(* IEC 61131-3 sources: PortalRobot/Portal_robot/Device/application/FB/FB_CELL_MANAGER (part 2) *)

(* ---- FB_CELL_MANAGER.CanReturnHeldBlank.st ---- *)
METHOD PRIVATE CanReturnHeldBlank : BOOL
VAR
	uiMagazine : UINT; // Магазин следующей операции, независимо от магазина возврата
	uiMachine  : UINT;
	uiType     : UINT;
	uiReservedFreeSlots : UINT; // Возврат занимает один универсальный слот своего магазина
END_VAR

// --- BEGIN IMPLEMENTATION ---

CanReturnHeldBlank := FALSE;

// Для одного типа возврат не открывает нового маршрута. Два груза сначала
// разбираются штатным LOAD/PUT; занятый исправный станок своей заготовки ждём.
IF (Config.uiTypeCount > UINT#1)
AND (Config.uiTypeCount <= UINT#3)
AND stRobotStatus.xBlankAvailable
AND NOT stRobotStatus.xDetailAvailable
AND NOT stRobotStatus.xBusy
AND NOT xStopRequested
AND xMagazineReady
AND (uiBlankPayloadType >= UINT#1)
AND (uiBlankPayloadType <= Config.uiTypeCount) THEN
	IF (stMagazineStatus.stTypeStatus.aiFreeSlot[uiBlankPayloadType] > SINT#0)
	AND (SelectMachineForHeldBlank(
		uiProductType := uiBlankPayloadType,
		uiCurrentMachine := uiSelectedMachine
	) = UINT#0) THEN
		FOR uiMagazine := UINT#1 TO GVL_CELL_SETTINGS.MagazineCount DO
			IF ((uiMagazine = UINT#1) AND xMagazine1Available)
			OR ((uiMagazine = UINT#2) AND xMagazine2Available) THEN
				uiReservedFreeSlots := UINT#0;
				IF uiMagazine = uiActiveMagazine THEN
					uiReservedFreeSlots := UINT#1;
				END_IF;
				FOR uiMachine := FIRST_MACHINE TO LAST_MACHINE DO
					IF IsMachineEligible(uiMachine := uiMachine) THEN
						uiType := Config.auiMachineType[uiMachine];
						IF uiType <> uiBlankPayloadType THEN
							// TAKE освобождает место даже в полной палете. Работающий
							// станок другого типа допускает обычное ожидание его цикла.
							IF (astMagazineStatus[uiMagazine].stTypeStatus.aiBlankSlot[uiType] > SINT#0)
							AND (astMachineStatus[uiMachine].xProcessing
								OR axMachineStartPending[uiMachine]
								OR (astMachineStatus[uiMachine].xCanAcceptService
									AND ((astMachineStatus[uiMachine].ePartState = E_PART_STATE.EMPTY)
										OR astMachineStatus[uiMachine].xServiceRequired))) THEN
								CanReturnHeldBlank := TRUE;
							END_IF;
							// Отдельная выгрузка полезна только для уже готовой детали.
							// Последний свободный слот нельзя занять возвратом и затем
							// выдать UNLOAD без места для этой детали.
							IF astMachineStatus[uiMachine].xCanAcceptService
							AND astMachineStatus[uiMachine].xServiceRequired
							AND (astMachineStatus[uiMachine].ePartState = E_PART_STATE.LOADED)
							AND (astMachineStatus[uiMachine].ePartType = E_PART_TYPE.DETAIL)
							AND (astMagazineStatus[uiMagazine].stTypeStatus.auiFreeCount[uiType] > uiReservedFreeSlots) THEN
								CanReturnHeldBlank := TRUE;
							END_IF;
						END_IF;
					END_IF;
				END_FOR;
			END_IF;
		END_FOR;
	END_IF;
END_IF;

(* ---- FB_CELL_MANAGER.HasMagazineWork.st ---- *)
METHOD PRIVATE HasMagazineWork : BOOL
VAR_INPUT
	uiMagazine : UINT; // Оцениваемый магазин; активный владелец не меняется
	xSupplyBlankOnly : BOOL; // TRUE: нужна именно допустимая подача заготовки
END_VAR
VAR
	uiMachine : UINT;
	uiType : UINT;
	xPending : BOOL;
END_VAR

// --- BEGIN IMPLEMENTATION ---

HasMagazineWork := FALSE;
IF (uiMagazine >= UINT#1) AND (uiMagazine <= UINT#2) THEN
	FOR uiMachine := FIRST_MACHINE TO LAST_MACHINE DO
		IF IsMachineEligible(uiMachine := uiMachine) THEN
			uiType := Config.auiMachineType[uiMachine];
			IF (uiType >= UINT#1) AND (uiType <= UINT#3) THEN
				xPending := IsMachineWorkPending(uiMachine := uiMachine);
				// Те же критерии, что у SelectMachineBeforeTake: готовый
				// LOAD/CHANGE либо ожидаемое автоматическое обслуживание.
				IF (astMagazineStatus[uiMagazine].stTypeStatus.aiBlankSlot[uiType] > SINT#0)
				AND (xPending OR (astMachineStatus[uiMachine].xCanAcceptService
					AND ((astMachineStatus[uiMachine].ePartState = E_PART_STATE.EMPTY)
						OR astMachineStatus[uiMachine].xServiceRequired))) THEN
					HasMagazineWork := TRUE;
				END_IF;
				// Без заготовки остаётся отдельный UNLOAD в свободный слот.
				IF NOT xSupplyBlankOnly
				AND (astMagazineStatus[uiMagazine].stTypeStatus.aiFreeSlot[uiType] > SINT#0)
				AND (xPending OR (astMachineStatus[uiMachine].xCanAcceptService
					AND astMachineStatus[uiMachine].xServiceRequired
					AND (astMachineStatus[uiMachine].ePartState = E_PART_STATE.LOADED)
					AND (astMachineStatus[uiMachine].ePartType = E_PART_TYPE.DETAIL))) THEN
					HasMagazineWork := TRUE;
				END_IF;
			END_IF;
		END_IF;
	END_FOR;
END_IF;

(* ---- FB_CELL_MANAGER.IsMachineCompatible.st ---- *)
METHOD PRIVATE IsMachineCompatible : BOOL
VAR_INPUT
	uiMachine     : UINT; // Проверяемый станок
	uiProductType : UINT; // Тип заготовки в захвате
END_VAR

// --- BEGIN IMPLEMENTATION ---

IsMachineCompatible := IsMachineEligible(uiMachine := uiMachine);
IF IsMachineCompatible THEN
	IsMachineCompatible := (uiProductType >= UINT#1)
		AND (uiProductType <= Config.uiTypeCount)
		AND (Config.auiMachineType[uiMachine] = uiProductType);
END_IF;

(* ---- FB_CELL_MANAGER.IsMachineEligible.st ---- *)
METHOD PRIVATE IsMachineEligible : BOOL
VAR_INPUT
	uiMachine : UINT; // Проверяемый станок
END_VAR

// --- BEGIN IMPLEMENTATION ---

IsMachineEligible := (uiMachine >= FIRST_MACHINE)
	AND (uiMachine <= LAST_MACHINE);

IF IsMachineEligible THEN
	IsMachineEligible := astMachineStatus[uiMachine].xEnabled
		AND NOT astMachineStatus[uiMachine].xError
		AND NOT astMachineStatus[uiMachine].xDisablePending
		AND NOT axGeometryUnloadBlocked[uiMachine]
		AND (Config.auiMachineType[uiMachine] >= UINT#1)
		AND (Config.auiMachineType[uiMachine] <= Config.uiTypeCount);
END_IF;

(* ---- FB_CELL_MANAGER.IsMachineWorkPending.st ---- *)
METHOD PRIVATE IsMachineWorkPending : BOOL
VAR_INPUT
	uiMachine : UINT; // Проверяемый станок
END_VAR

// --- BEGIN IMPLEMENTATION ---

IsMachineWorkPending := FALSE;
IF IsMachineEligible(uiMachine := uiMachine) THEN
	// LOADED сам по себе не обещает автоматического продолжения: оператор
	// может ещё не разрешить цикл. Сохраняем обработку, подтверждение запуска
	// и короткий автоматический переход после обработки/обслуживания.
	IsMachineWorkPending := astMachineStatus[uiMachine].xProcessing
		OR axMachineStartPending[uiMachine]
		OR ((astMachineStatus[uiMachine].ePartState = E_PART_STATE.LOADED)
			AND ((astMachineStatus[uiMachine].ePartType = E_PART_TYPE.PART)
				OR (astMachineStatus[uiMachine].ePartType = E_PART_TYPE.DETAIL))
			AND (astMachineStatus[uiMachine].xBusy
				OR astMachineStatus[uiMachine].xDone));
END_IF;

(* ---- FB_CELL_MANAGER.PlanGeometry.st ---- *)
METHOD PRIVATE PlanGeometry : BOOL
VAR
	uiFree : UINT;
	uiAvailable : UINT;
END_VAR

// --- BEGIN IMPLEMENTATION ---

PlanGeometry := FALSE;
IF xGeometryHeld AND stRobotStatus.xDetailAvailable AND (uiGeometryMachine >= UINT#1) AND (uiGeometryMachine <= UINT#3) THEN
	uiFree := F_GEOMETRY_SELECT_STATION(xRequireFree := TRUE, uiMachine := uiGeometryMachine);
	uiAvailable := F_GEOMETRY_SELECT_STATION(xRequireFree := FALSE, uiMachine := uiGeometryMachine);
	IF uiFree > UINT#0 THEN
		uiGeometryStation := uiFree; uiGeometryStep := UINT#0;
		GVL_GEOMETRY_CONTROL.astCalls[uiGeometryMachine].uiStation := uiFree;
		GVL_GEOMETRY_CONTROL.astCalls[uiGeometryMachine].uiState := UINT#3;
		GVL_GEOMETRY_CONTROL.astCalls[uiGeometryMachine].uiReason := UINT#0;
		F_GEOMETRY_EVENT(Call := GVL_GEOMETRY_CONTROL.astCalls[uiGeometryMachine]);
		GVL_GEOMETRY_CONTROL.astSignals[uiFree].Call := GVL_GEOMETRY_CONTROL.astCalls[uiGeometryMachine];
		GVL_GEOMETRY_CONTROL.astSignals[uiFree].xReserve := TRUE;
		eState := E_CELL_MANAGER_STATE.GEOMETRY_DELIVER; PlanGeometry := TRUE;
	ELSIF (uiAvailable > UINT#0) AND Persistent_Value.xWaitWhenOccupied THEN
		uiGeometryParkStation := uiAvailable;
		eState := E_CELL_MANAGER_STATE.GEOMETRY_WAIT_FREE; PlanGeometry := TRUE;
	ELSE
		// Окончательный журнал магазина формируем только по фактической укладке.
		IF uiAvailable > UINT#0 THEN uiGeometryBypassReason := UINT#1; ELSE uiGeometryBypassReason := UINT#2; END_IF;
		udiGeometryMagazineCounter := stMagazineStatus.udiProducedPartsTotal;
	END_IF;
END_IF;

(* ---- FB_CELL_MANAGER.RaisePayloadRouteWarning.st ---- *)
METHOD PRIVATE RaisePayloadRouteWarning
VAR_INPUT
	uiPayloadType     : UINT;
	uiDestinationType : UINT;
END_VAR

// --- BEGIN IMPLEMENTATION ---

IF (uiPayloadType >= UINT#1)
AND (uiDestinationType >= UINT#1)
AND (uiPayloadType <> uiDestinationType) THEN
	IF NOT xPayloadRouteWarningActive THEN
		Diag.stWarning.uiCode := WRN_PAYLOAD_ROUTE_MISMATCH;
		Diag.stWarning.udiSequence := Diag.stWarning.udiSequence + UDINT#1;
		IF Diag.stWarning.udiSequence = UDINT#0 THEN
			Diag.stWarning.udiSequence := UDINT#1;
		END_IF;
		xPayloadRouteWarningActive := TRUE;
	END_IF;
ELSE
	xPayloadRouteWarningActive := FALSE;
END_IF;

(* ---- FB_CELL_MANAGER.RunGeometryRoute.st ---- *)
METHOD PRIVATE RunGeometryRoute

// --- BEGIN IMPLEMENTATION ---

CASE eState OF
	E_CELL_MANAGER_STATE.GEOMETRY_WAIT_FREE:
		IF uiGeometryParkStation = UINT#1 THEN eGeometrySafePoint := E_POINT_NAME.GEOMETRY_1_SAFE;
		ELSE eGeometrySafePoint := E_POINT_NAME.GEOMETRY_2_SAFE; END_IF;
		IF stRobotStatus.xBusy OR stRobotStatus.xDone OR xMotionBusy THEN
			// Освобождение ГК не отменяет уже выданное парковочное движение.
			Command.stRobot.xExecute := TRUE; Command.stRobot.eAction := E_ROBOT_ACTION.MOVE_TO_POINT;
			Command.stRobot.eSetPoint := eGeometrySafePoint;
			IF stRobotStatus.xDone THEN eGeometryReturnState := E_CELL_MANAGER_STATE.GEOMETRY_WAIT_FREE; eState := E_CELL_MANAGER_STATE.GEOMETRY_RELEASE_COMMAND; END_IF;
		ELSIF xStopRequested THEN
			xRunning := FALSE; eState := E_CELL_MANAGER_STATE.IDLE;
		ELSIF F_GEOMETRY_SELECT_STATION(xRequireFree := TRUE, uiMachine := uiGeometryMachine) > UINT#0 THEN
			eState := E_CELL_MANAGER_STATE.PLAN_TARGET;
		ELSIF (F_GEOMETRY_SELECT_STATION(xRequireFree := FALSE, uiMachine := uiGeometryMachine) = UINT#0) OR NOT Persistent_Value.xWaitWhenOccupied THEN
			eState := E_CELL_MANAGER_STATE.PLAN_TARGET;
		ELSE
			// Ожидаем с деталью в захвате на безопасной высоте; конвейер может работать.
			IF uiGeometryParkStation = UINT#1 THEN eGeometrySafePoint := E_POINT_NAME.GEOMETRY_1_SAFE;
			ELSE eGeometrySafePoint := E_POINT_NAME.GEOMETRY_2_SAFE; END_IF;
			IF stRobotStatus.eCurrentPoint <> eGeometrySafePoint THEN
				Command.stRobot.xExecute := TRUE; Command.stRobot.eAction := E_ROBOT_ACTION.MOVE_TO_POINT;
				Command.stRobot.eSetPoint := eGeometrySafePoint;
				IF stRobotStatus.xDone THEN eGeometryReturnState := E_CELL_MANAGER_STATE.GEOMETRY_WAIT_FREE; eState := E_CELL_MANAGER_STATE.GEOMETRY_RELEASE_COMMAND; END_IF;
			END_IF;
		END_IF;
	E_CELL_MANAGER_STATE.GEOMETRY_DELIVER:
		IF (uiGeometryStation < UINT#1) OR (uiGeometryStation > UINT#2) THEN
			Error.dwErrorActive := Error.dwErrorActive OR ERR_ROBOT; eState := E_CELL_MANAGER_STATE.ERROR;
		ELSIF GVL_GEOMETRY_CONTROL.astStatus[uiGeometryStation].xError
		AND NOT GVL_GEOMETRY_CONTROL.astSignals[uiGeometryStation].xRobotInteraction THEN
			// Оборудование отказало до входа: робот может выбрать другой ГК.
			GVL_GEOMETRY_CONTROL.astSignals[uiGeometryStation].xReserve := FALSE;
			GVL_GEOMETRY_CONTROL.astSignals[uiGeometryStation].xReleased := TRUE;
			GVL_GEOMETRY_CONTROL.astCalls[uiGeometryMachine].uiStation := UINT#0;
			GVL_GEOMETRY_CONTROL.astCalls[uiGeometryMachine].uiState := UINT#2;
			GVL_GEOMETRY_CONTROL.astCalls[uiGeometryMachine].uiReason := UINT#4;
			F_GEOMETRY_EVENT(Call := GVL_GEOMETRY_CONTROL.astCalls[uiGeometryMachine]);
			uiGeometryStation := UINT#0; eState := E_CELL_MANAGER_STATE.PLAN_TARGET;
		ELSIF NOT GVL_GEOMETRY_CONTROL.astSignals[uiGeometryStation].xRobotInteraction
		AND (NOT GVL_GEOMETRY_CONTROL.astStatus[uiGeometryStation].xEnabled
			OR (GVL_GEOMETRY_CONTROL.astStatus[uiGeometryStation].uiState = UINT#5)
			OR GVL_GEOMETRY_CONTROL.astStatus[uiGeometryStation].xDriveRunning) THEN
			// Выключение в том же скане, что резерв, не разрешает вход робота.
			GVL_GEOMETRY_CONTROL.astSignals[uiGeometryStation].xReserve := FALSE;
			GVL_GEOMETRY_CONTROL.astSignals[uiGeometryStation].xReleased := TRUE;
			GVL_GEOMETRY_CONTROL.astCalls[uiGeometryMachine].uiStation := UINT#0;
			GVL_GEOMETRY_CONTROL.astCalls[uiGeometryMachine].uiState := UINT#2;
			GVL_GEOMETRY_CONTROL.astCalls[uiGeometryMachine].uiReason := UINT#3;
			F_GEOMETRY_EVENT(Call := GVL_GEOMETRY_CONTROL.astCalls[uiGeometryMachine]);
			uiGeometryStation := UINT#0; eState := E_CELL_MANAGER_STATE.PLAN_TARGET;
		ELSIF GVL_GEOMETRY_CONTROL.astStatus[uiGeometryStation].xError OR stRobotStatus.xError OR xGlobalError THEN
			xSafetyHomeRequired := TRUE; xStoppedPoseValid := FALSE;
			Error.dwErrorActive := Error.dwErrorActive OR ERR_ROBOT; eState := E_CELL_MANAGER_STATE.ERROR;
		ELSIF GVL_GEOMETRY_CONTROL.astStatus[uiGeometryStation].xReserved THEN
			IF uiGeometryStation = UINT#1 THEN
				eGeometrySafePoint := E_POINT_NAME.GEOMETRY_1_SAFE; eGeometryPlacePoint := E_POINT_NAME.GEOMETRY_1_PLACE;
			ELSE
				eGeometrySafePoint := E_POINT_NAME.GEOMETRY_2_SAFE; eGeometryPlacePoint := E_POINT_NAME.GEOMETRY_2_PLACE;
			END_IF;
			GVL_GEOMETRY_CONTROL.astSignals[uiGeometryStation].xRobotInteraction := TRUE;
			IF uiGeometryStep <= UINT#4 THEN
				Command.stRobot.xExecute := TRUE; Command.stRobot.eAction := E_ROBOT_ACTION.MOVE_TO_POINT;
				CASE uiGeometryStep OF
					UINT#0, UINT#4: Command.stRobot.eSetPoint := eGeometrySafePoint;
					// Для укладки на ГК нужна ориентация «к заготовке»; поворот выполняется на SAFE.
					UINT#1: Command.stRobot.eAction := E_ROBOT_ACTION.ROTATE_TO_BLANK;
					UINT#2: Command.stRobot.eSetPoint := eGeometryPlacePoint;
					UINT#3: Command.stRobot.eAction := E_ROBOT_ACTION.UNCLAMP_2;
				END_CASE;
				IF stRobotStatus.xDone THEN
					IF uiGeometryStep = UINT#3 THEN
						IF stRobotStatus.xGripper2Open AND NOT stRobotStatus.xDetailAvailable THEN
							GVL_GEOMETRY_CONTROL.astSignals[uiGeometryStation].xDeposited := TRUE;
							uiDetailPayloadType := UINT#0;
						ELSE Error.dwErrorActive := Error.dwErrorActive OR ERR_ROBOT; eState := E_CELL_MANAGER_STATE.ERROR; END_IF;
					END_IF;
					IF eState <> E_CELL_MANAGER_STATE.ERROR THEN
						eGeometryReturnState := E_CELL_MANAGER_STATE.GEOMETRY_DELIVER;
						eState := E_CELL_MANAGER_STATE.GEOMETRY_RELEASE_COMMAND;
					END_IF;
				END_IF;
			ELSE
				GVL_GEOMETRY_CONTROL.astSignals[uiGeometryStation].xReserve := FALSE;
				GVL_GEOMETRY_CONTROL.astSignals[uiGeometryStation].xDeposited := FALSE;
				GVL_GEOMETRY_CONTROL.astSignals[uiGeometryStation].xRobotInteraction := FALSE;
				GVL_GEOMETRY_CONTROL.astSignals[uiGeometryStation].xReleased := TRUE;
				GVL_GEOMETRY_CONTROL.uiLastStation := uiGeometryStation;
				xGeometryHeld := FALSE; uiGeometryMachine := UINT#0; uiGeometryStation := UINT#0;
				eState := E_CELL_MANAGER_STATE.PLAN_TARGET;
			END_IF;
		ELSE
			// Потеря резерва в зоне робота требует восстановления, а не нового маршрута.
			IF GVL_GEOMETRY_CONTROL.astSignals[uiGeometryStation].xRobotInteraction THEN
				xSafetyHomeRequired := TRUE; xStoppedPoseValid := FALSE;
				Error.dwErrorActive := Error.dwErrorActive OR ERR_ROBOT; eState := E_CELL_MANAGER_STATE.ERROR;
			ELSIF NOT GVL_GEOMETRY_CONTROL.astStatus[uiGeometryStation].xReady
			OR (GVL_GEOMETRY_CONTROL.astStatus[uiGeometryStation].uiState = UINT#5) THEN
				GVL_GEOMETRY_CONTROL.astSignals[uiGeometryStation].xReserve := FALSE;
				GVL_GEOMETRY_CONTROL.astSignals[uiGeometryStation].xReleased := TRUE;
				GVL_GEOMETRY_CONTROL.astCalls[uiGeometryMachine].uiStation := UINT#0;
				GVL_GEOMETRY_CONTROL.astCalls[uiGeometryMachine].uiState := UINT#2;
				GVL_GEOMETRY_CONTROL.astCalls[uiGeometryMachine].uiReason := UINT#3;
				F_GEOMETRY_EVENT(Call := GVL_GEOMETRY_CONTROL.astCalls[uiGeometryMachine]);
				uiGeometryStation := UINT#0; eState := E_CELL_MANAGER_STATE.PLAN_TARGET;
			END_IF;
		END_IF;
	E_CELL_MANAGER_STATE.GEOMETRY_RELEASE_COMMAND:
		IF stRobotStatus.xError THEN
			xSafetyHomeRequired := TRUE; xStoppedPoseValid := FALSE;
			Error.dwErrorActive := Error.dwErrorActive OR ERR_ROBOT; eState := E_CELL_MANAGER_STATE.ERROR;
		ELSIF NOT stRobotStatus.xBusy AND NOT stRobotStatus.xDone THEN
			IF eGeometryReturnState = E_CELL_MANAGER_STATE.GEOMETRY_DELIVER THEN uiGeometryStep := uiGeometryStep + UINT#1; END_IF;
			eState := eGeometryReturnState;
		END_IF;
END_CASE;

(* ---- FB_CELL_MANAGER.SelectMachineBeforeTake.st ---- *)
METHOD PRIVATE SelectMachineBeforeTake : UINT
VAR
	uiMachine           : UINT; // Проверяемый станок
	uiType              : UINT; // Тип станка
	xTimedFound         : BOOL; // Найден кандидат с оценкой времени
	tMinimumRemaining   : TIME; // Минимальное найденное оставшееся время
	tCandidateRemaining : TIME; // Оценка кандидата, который подтверждает запуск цикла
END_VAR

// --- BEGIN IMPLEMENTATION ---

SelectMachineBeforeTake := UINT#0;
xTimedFound := FALSE;
tMinimumRemaining := T#0S;

// Сначала выбирается станок, который можно обслужить без ожидания.
// xPartReady отдельно не используется: после завершения обслуживания он может
// сохраняться до перехода FB_MACHINE из DONE в IDLE и повторно выбрать тот же станок.
FOR uiMachine := FIRST_MACHINE TO LAST_MACHINE DO
	uiType := Config.auiMachineType[uiMachine];
	IF IsMachineEligible(uiMachine := uiMachine) THEN
		IF (SelectMachineBeforeTake = UINT#0)
		AND (stMagazineStatus.stTypeStatus.aiBlankSlot[uiType] > SINT#0)
		AND astMachineStatus[uiMachine].xCanAcceptService
		AND ((astMachineStatus[uiMachine].ePartState = E_PART_STATE.EMPTY)
			OR astMachineStatus[uiMachine].xServiceRequired) THEN
			SelectMachineBeforeTake := uiMachine;
		END_IF;
	END_IF;
END_FOR;

// Затем сравниваются фактически обрабатывающие станки по оставшемуся времени.
IF SelectMachineBeforeTake = UINT#0 THEN
	FOR uiMachine := FIRST_MACHINE TO LAST_MACHINE DO
		uiType := Config.auiMachineType[uiMachine];
		IF IsMachineEligible(uiMachine := uiMachine) THEN
			IF (stMagazineStatus.stTypeStatus.aiBlankSlot[uiType] > SINT#0)
			AND astMachineStatus[uiMachine].xProcessing
			AND astMachineStatus[uiMachine].xCycleTimeValid THEN
				IF NOT xTimedFound
				OR (astMachineStatus[uiMachine].tRemaining < tMinimumRemaining) THEN
					SelectMachineBeforeTake := uiMachine;
					tMinimumRemaining := astMachineStatus[uiMachine].tRemaining;
					xTimedFound := TRUE;
				END_IF;
			END_IF;
		END_IF;
	END_FOR;
END_IF;

// Только что обслуженный станок может появиться в xProcessing на несколько циклов PLC позже.
// До подтверждения запуска он участвует в том же сравнении по полному tCycleExpected.
IF (SelectMachineBeforeTake = UINT#0) OR xTimedFound THEN
	FOR uiMachine := FIRST_MACHINE TO LAST_MACHINE DO
		uiType := Config.auiMachineType[uiMachine];
		IF axMachineStartPending[uiMachine]
		AND IsMachineEligible(uiMachine := uiMachine)
		AND (stMagazineStatus.stTypeStatus.aiBlankSlot[uiType] > SINT#0)
		AND astMachineStatus[uiMachine].xCycleTimeValid THEN
			tCandidateRemaining := START_PENDING_ESTIMATE
				+ astMachineStatus[uiMachine].tCycleExpected;
			IF NOT xTimedFound
			OR (tCandidateRemaining < tMinimumRemaining) THEN
				SelectMachineBeforeTake := uiMachine;
				tMinimumRemaining := tCandidateRemaining;
				xTimedFound := TRUE;
			END_IF;
		END_IF;
	END_FOR;
END_IF;

// Неизвестное время не делает включённый исправный станок недоступным.
IF (SelectMachineBeforeTake = UINT#0) AND NOT xTimedFound THEN
	FOR uiMachine := FIRST_MACHINE TO LAST_MACHINE DO
		uiType := Config.auiMachineType[uiMachine];
		IF IsMachineEligible(uiMachine := uiMachine) THEN
			IF (SelectMachineBeforeTake = UINT#0)
			AND (stMagazineStatus.stTypeStatus.aiBlankSlot[uiType] > SINT#0)
			AND IsMachineWorkPending(uiMachine := uiMachine) THEN
				SelectMachineBeforeTake := uiMachine;
			END_IF;
		END_IF;
	END_FOR;
END_IF;

(* ---- FB_CELL_MANAGER.SelectMachineForHeldBlank.st ---- *)
METHOD PRIVATE SelectMachineForHeldBlank : UINT
VAR_INPUT
	uiProductType    : UINT; // Тип уже взятой заготовки
	uiCurrentMachine : UINT; // Текущая цель для устойчивого повторного выбора
END_VAR
VAR
	uiMachine           : UINT; // Проверяемый станок
	xTimedFound         : BOOL; // Найден станок с оценкой времени
	xCurrentTimed       : BOOL; // Текущая цель имеет сопоставимую оценку
	tMinimumRemaining   : TIME; // Минимальное оставшееся время
	tCandidateRemaining : TIME; // Оценка проверяемого станка
	tCurrentRemaining   : TIME; // Оценка текущей цели
END_VAR

// --- BEGIN IMPLEMENTATION ---

SelectMachineForHeldBlank := UINT#0;
xTimedFound := FALSE;
xCurrentTimed := FALSE;
tMinimumRemaining := T#0S;
tCandidateRemaining := T#0S;
tCurrentRemaining := T#0S;

// UINT#0 означает, что после остановки/аварии текущая цель ещё не выбрана.
// Проверка диапазона вынесена отдельно: обычный AND в CODESYS вычисляет все
// операнды и не защищает ARRAY [1..3] от обращения по индексу 0.
IF (uiCurrentMachine >= FIRST_MACHINE)
AND (uiCurrentMachine <= LAST_MACHINE) THEN
	// Если робот уже находится у готовой совместимой цели, лишнее перемещение не требуется.
	IF IsMachineCompatible(
		uiMachine := uiCurrentMachine,
		uiProductType := uiProductType
	)
	AND astMachineStatus[uiCurrentMachine].xCanAcceptService
	AND ((astMachineStatus[uiCurrentMachine].ePartState = E_PART_STATE.EMPTY)
		OR astMachineStatus[uiCurrentMachine].xServiceRequired) THEN
		SelectMachineForHeldBlank := uiCurrentMachine;
	END_IF;
END_IF;

// Готовая совместимая цель имеет приоритет. Переходный xPartReady без
// xCanAcceptService не считается разрешением на повторное обслуживание.
FOR uiMachine := FIRST_MACHINE TO LAST_MACHINE DO
	IF (SelectMachineForHeldBlank = UINT#0)
	AND IsMachineEligible(uiMachine := uiMachine)
	AND (Config.auiMachineType[uiMachine] = uiProductType)
	AND astMachineStatus[uiMachine].xCanAcceptService
	AND ((astMachineStatus[uiMachine].ePartState = E_PART_STATE.EMPTY)
		OR astMachineStatus[uiMachine].xServiceRequired) THEN
		SelectMachineForHeldBlank := uiMachine;
	END_IF;
END_FOR;

// Обрабатывающие и только что запущенные совместимые станки сравниваются
// по одному прогнозу: tRemaining либо полный tCycleExpected для start-pending.
IF SelectMachineForHeldBlank = UINT#0 THEN
	FOR uiMachine := FIRST_MACHINE TO LAST_MACHINE DO
		IF IsMachineEligible(uiMachine := uiMachine)
		AND (Config.auiMachineType[uiMachine] = uiProductType)
		AND astMachineStatus[uiMachine].xCycleTimeValid THEN
			IF astMachineStatus[uiMachine].xProcessing THEN
				tCandidateRemaining := astMachineStatus[uiMachine].tRemaining;
			ELSIF axMachineStartPending[uiMachine] THEN
				tCandidateRemaining := START_PENDING_ESTIMATE
					+ astMachineStatus[uiMachine].tCycleExpected;
			ELSE
				tCandidateRemaining := T#0S;
			END_IF;

			IF astMachineStatus[uiMachine].xProcessing
			OR axMachineStartPending[uiMachine] THEN
				IF NOT xTimedFound
				OR (tCandidateRemaining < tMinimumRemaining) THEN
					SelectMachineForHeldBlank := uiMachine;
					tMinimumRemaining := tCandidateRemaining;
					xTimedFound := TRUE;
				END_IF;
			END_IF;
		END_IF;
	END_FOR;

	// При почти одинаковом времени сохраняется текущая цель.
	IF xTimedFound
	AND (uiCurrentMachine >= FIRST_MACHINE)
	AND (uiCurrentMachine <= LAST_MACHINE) THEN
		IF (SelectMachineForHeldBlank <> uiCurrentMachine)
		AND IsMachineCompatible(
			uiMachine := uiCurrentMachine,
			uiProductType := uiProductType
		)
		AND astMachineStatus[uiCurrentMachine].xCycleTimeValid THEN
			xCurrentTimed := astMachineStatus[uiCurrentMachine].xProcessing
				OR axMachineStartPending[uiCurrentMachine];
			IF astMachineStatus[uiCurrentMachine].xProcessing THEN
				tCurrentRemaining := astMachineStatus[uiCurrentMachine].tRemaining;
			ELSIF axMachineStartPending[uiCurrentMachine] THEN
				tCurrentRemaining := START_PENDING_ESTIMATE
					+ astMachineStatus[uiCurrentMachine].tCycleExpected;
			END_IF;
			IF xCurrentTimed
			AND (tCurrentRemaining >= tMinimumRemaining)
			AND ((tCurrentRemaining - tMinimumRemaining) <= MACHINE_SWITCH_DEADBAND) THEN
				SelectMachineForHeldBlank := uiCurrentMachine;
			END_IF;
		END_IF;
	END_IF;
END_IF;

// Без точной оценки сохраняется текущий обрабатывающий маршрут либо выбирается
// первый совместимый обрабатывающий/start-pending станок.
IF SelectMachineForHeldBlank = UINT#0 THEN
	IF (uiCurrentMachine >= FIRST_MACHINE)
	AND (uiCurrentMachine <= LAST_MACHINE) THEN
		IF IsMachineCompatible(
			uiMachine := uiCurrentMachine,
			uiProductType := uiProductType
		)
		AND (astMachineStatus[uiCurrentMachine].xProcessing
			OR axMachineStartPending[uiCurrentMachine]) THEN
			SelectMachineForHeldBlank := uiCurrentMachine;
		END_IF;
	END_IF;

	FOR uiMachine := FIRST_MACHINE TO LAST_MACHINE DO
		IF (SelectMachineForHeldBlank = UINT#0)
		AND IsMachineEligible(uiMachine := uiMachine)
		AND (Config.auiMachineType[uiMachine] = uiProductType)
		AND (astMachineStatus[uiMachine].xProcessing
			OR axMachineStartPending[uiMachine]) THEN
			SelectMachineForHeldBlank := uiMachine;
		END_IF;
	END_FOR;
END_IF;

// Включённая исправная цель сохраняет ожидание своей заготовки, даже если
// станок ещё не готов. Нулевой результат только разрешает проверку полезности
// возврата в SELECT_FALLBACK; сам по себе он не требует RETURN_BLANK.
IF SelectMachineForHeldBlank = UINT#0 THEN
	IF (uiCurrentMachine >= FIRST_MACHINE)
	AND (uiCurrentMachine <= LAST_MACHINE) THEN
		IF IsMachineCompatible(
			uiMachine := uiCurrentMachine,
			uiProductType := uiProductType
		) THEN
			SelectMachineForHeldBlank := uiCurrentMachine;
		END_IF;
	END_IF;

	FOR uiMachine := FIRST_MACHINE TO LAST_MACHINE DO
		IF (SelectMachineForHeldBlank = UINT#0)
		AND IsMachineEligible(uiMachine := uiMachine)
		AND (Config.auiMachineType[uiMachine] = uiProductType) THEN
			SelectMachineForHeldBlank := uiMachine;
		END_IF;
	END_FOR;
END_IF;

(* ---- FB_CELL_MANAGER.SelectMachineForUnload.st ---- *)
METHOD PRIVATE SelectMachineForUnload : UINT
VAR_INPUT
	uiCurrentMachine : UINT; // Текущая цель для устойчивого повторного выбора
END_VAR
VAR
	uiMachine           : UINT; // Проверяемый станок
	uiType              : UINT; // Тип детали станка
	xTimedFound         : BOOL; // Найден станок с оценкой времени
	xCurrentTimed       : BOOL; // Текущая цель имеет сопоставимую оценку
	tMinimumRemaining   : TIME; // Минимальное найденное оставшееся время
	tCandidateRemaining : TIME; // Оценка проверяемого станка
	tCurrentRemaining   : TIME; // Оценка текущей цели
END_VAR

// --- BEGIN IMPLEMENTATION ---

SelectMachineForUnload := UINT#0;
xTimedFound := FALSE;
xCurrentTimed := FALSE;
tMinimumRemaining := T#0S;
tCandidateRemaining := T#0S;
tCurrentRemaining := T#0S;

// Если робот уже ждёт над готовым станком, лишнее перемещение не требуется.
IF (uiCurrentMachine >= FIRST_MACHINE)
AND (uiCurrentMachine <= LAST_MACHINE) THEN
	IF IsMachineEligible(uiMachine := uiCurrentMachine) THEN
		uiType := Config.auiMachineType[uiCurrentMachine];
		IF (stMagazineStatus.stTypeStatus.aiFreeSlot[uiType] > SINT#0)
		AND astMachineStatus[uiCurrentMachine].xCanAcceptService
		AND astMachineStatus[uiCurrentMachine].xServiceRequired
		AND (astMachineStatus[uiCurrentMachine].ePartState = E_PART_STATE.LOADED)
		AND (astMachineStatus[uiCurrentMachine].ePartType = E_PART_TYPE.DETAIL) THEN
			SelectMachineForUnload := uiCurrentMachine;
		END_IF;
	END_IF;
END_IF;

// Готовая деталь имеет приоритет над ожиданием обработки.
FOR uiMachine := FIRST_MACHINE TO LAST_MACHINE DO
	uiType := Config.auiMachineType[uiMachine];
	IF IsMachineEligible(uiMachine := uiMachine) THEN
		IF (SelectMachineForUnload = UINT#0)
		AND astMachineStatus[uiMachine].xCanAcceptService
		AND astMachineStatus[uiMachine].xServiceRequired
		AND (astMachineStatus[uiMachine].ePartState = E_PART_STATE.LOADED)
		AND (astMachineStatus[uiMachine].ePartType = E_PART_TYPE.DETAIL)
		AND (stMagazineStatus.stTypeStatus.aiFreeSlot[uiType] > SINT#0) THEN
			SelectMachineForUnload := uiMachine;
		END_IF;
	END_IF;
END_FOR;

// Если готовых деталей пока нет, робот заранее направляется к станку с
// минимальным оставшимся временем обработки.
IF SelectMachineForUnload = UINT#0 THEN
	FOR uiMachine := FIRST_MACHINE TO LAST_MACHINE DO
		uiType := Config.auiMachineType[uiMachine];
		IF IsMachineEligible(uiMachine := uiMachine) THEN
			IF (stMagazineStatus.stTypeStatus.aiFreeSlot[uiType] > SINT#0)
			AND astMachineStatus[uiMachine].xCycleTimeValid THEN
				IF astMachineStatus[uiMachine].xProcessing THEN
					tCandidateRemaining := astMachineStatus[uiMachine].tRemaining;
				ELSIF axMachineStartPending[uiMachine] THEN
					tCandidateRemaining := START_PENDING_ESTIMATE
						+ astMachineStatus[uiMachine].tCycleExpected;
				ELSE
					tCandidateRemaining := T#0S;
				END_IF;

				IF astMachineStatus[uiMachine].xProcessing
				OR axMachineStartPending[uiMachine] THEN
					IF NOT xTimedFound
					OR (tCandidateRemaining < tMinimumRemaining) THEN
						SelectMachineForUnload := uiMachine;
						tMinimumRemaining := tCandidateRemaining;
						xTimedFound := TRUE;
					END_IF;
				END_IF;
			END_IF;
		END_IF;
	END_FOR;

	// При почти одинаковом времени сохраняется уже выбранная цель.
	IF xTimedFound
	AND (uiCurrentMachine >= FIRST_MACHINE)
	AND (uiCurrentMachine <= LAST_MACHINE) THEN
		IF (SelectMachineForUnload <> uiCurrentMachine)
		AND IsMachineEligible(uiMachine := uiCurrentMachine) THEN
			uiType := Config.auiMachineType[uiCurrentMachine];
			IF (stMagazineStatus.stTypeStatus.aiFreeSlot[uiType] > SINT#0)
			AND astMachineStatus[uiCurrentMachine].xCycleTimeValid THEN
				xCurrentTimed := astMachineStatus[uiCurrentMachine].xProcessing
					OR axMachineStartPending[uiCurrentMachine];
				IF astMachineStatus[uiCurrentMachine].xProcessing THEN
					tCurrentRemaining := astMachineStatus[uiCurrentMachine].tRemaining;
				ELSIF axMachineStartPending[uiCurrentMachine] THEN
					tCurrentRemaining := START_PENDING_ESTIMATE
						+ astMachineStatus[uiCurrentMachine].tCycleExpected;
				END_IF;
				IF xCurrentTimed
				AND (tCurrentRemaining >= tMinimumRemaining)
				AND ((tCurrentRemaining - tMinimumRemaining) <= MACHINE_SWITCH_DEADBAND) THEN
					SelectMachineForUnload := uiCurrentMachine;
				END_IF;
			END_IF;
		END_IF;
	END_IF;
END_IF;

// При неизвестном времени сохраняется текущая цель либо выбирается первый
// обрабатывающийся/только что запущенный станок с доступным слотом.
IF SelectMachineForUnload = UINT#0 THEN
	IF (uiCurrentMachine >= FIRST_MACHINE)
	AND (uiCurrentMachine <= LAST_MACHINE) THEN
		IF IsMachineEligible(uiMachine := uiCurrentMachine) THEN
			uiType := Config.auiMachineType[uiCurrentMachine];
			IF (stMagazineStatus.stTypeStatus.aiFreeSlot[uiType] > SINT#0)
			AND (astMachineStatus[uiCurrentMachine].xProcessing
				OR axMachineStartPending[uiCurrentMachine]) THEN
				SelectMachineForUnload := uiCurrentMachine;
			END_IF;
		END_IF;
	END_IF;

	FOR uiMachine := FIRST_MACHINE TO LAST_MACHINE DO
		uiType := Config.auiMachineType[uiMachine];
		IF IsMachineEligible(uiMachine := uiMachine) THEN
			IF (SelectMachineForUnload = UINT#0)
			AND (stMagazineStatus.stTypeStatus.aiFreeSlot[uiType] > SINT#0)
			AND (astMachineStatus[uiMachine].xProcessing
				OR axMachineStartPending[uiMachine]) THEN
				SelectMachineForUnload := uiMachine;
			END_IF;
		END_IF;
	END_FOR;
END_IF;

// Переход от окончания цикла к готовности двери может занять несколько сканов.
// В это время сохраняется автоматически продолжающий работу станок.
// Ожидание решения оператора при LOADED сюда не входит.
IF SelectMachineForUnload = UINT#0 THEN
	IF (uiCurrentMachine >= FIRST_MACHINE)
	AND (uiCurrentMachine <= LAST_MACHINE) THEN
		IF IsMachineEligible(uiMachine := uiCurrentMachine) THEN
			uiType := Config.auiMachineType[uiCurrentMachine];
			IF (stMagazineStatus.stTypeStatus.aiFreeSlot[uiType] > SINT#0)
			AND IsMachineWorkPending(uiMachine := uiCurrentMachine) THEN
				SelectMachineForUnload := uiCurrentMachine;
			END_IF;
		END_IF;
	END_IF;

	FOR uiMachine := FIRST_MACHINE TO LAST_MACHINE DO
		uiType := Config.auiMachineType[uiMachine];
		IF IsMachineEligible(uiMachine := uiMachine) THEN
			IF (SelectMachineForUnload = UINT#0)
			AND (stMagazineStatus.stTypeStatus.aiFreeSlot[uiType] > SINT#0)
			AND IsMachineWorkPending(uiMachine := uiMachine) THEN
				SelectMachineForUnload := uiMachine;
			END_IF;
		END_IF;
	END_FOR;
END_IF;

(* ---- FB_CELL_MANAGER.UpdateErrorView.st ---- *)
METHOD PRIVATE UpdateErrorView : ST_CELL_ERROR
VAR_INPUT
	dwError : DWORD; // Битовая маска ошибок нового менеджера
END_VAR
VAR
	stError : ST_CELL_ERROR; // Совместимое представление ошибок
END_VAR

// --- BEGIN IMPLEMENTATION ---

stError.BOTH_GRIPPERS_OCCUPIED := (dwError AND ERR_BOTH_GRIPPERS) <> DWORD#0;
stError.ROBOT_ERROR := (dwError AND ERR_ROBOT) <> DWORD#0;
stError.MAGAZINE_ERROR := (dwError AND ERR_MAGAZINE) <> DWORD#0;
stError.MACHINE_ERROR := (dwError AND ERR_MACHINE) <> DWORD#0;
stError.GLOBAL_STOP := (dwError AND ERR_GLOBAL_STOP) <> DWORD#0;
UpdateErrorView := stError;

(* ---- FB_CELL_MANAGER.UpdateGeometryWait.st ---- *)
METHOD PRIVATE UpdateGeometryWait
VAR
	uiMachine : UINT;
	uiFreeStation : UINT;
	uiCallState : UINT;
	xCalled : BOOL;
	xReadyDetail : BOOL;
	xWaiting : BOOL;
	xRaiseWarning : BOOL;
	Call : ST_GEOMETRY_CALL;
	EmptyCall : ST_GEOMETRY_CALL;
END_VAR

// --- BEGIN IMPLEMENTATION ---

uiFreeStation := F_GEOMETRY_SELECT_STATION(xRequireFree := TRUE, uiMachine := UINT#0);
xRaiseWarning := FALSE;
FOR uiMachine := FIRST_MACHINE TO LAST_MACHINE DO
	uiCallState := GVL_GEOMETRY_CONTROL.astCalls[uiMachine].uiState;
	xCalled := uiCallState = UINT#1;
	// Автовызов известен до выгрузки; счётчик меняется только при фактическом взятии.
	IF ((uiCallState = UINT#0) OR (uiCallState > UINT#3))
	AND GVL_GEOMETRY_CONTROL.xSupported AND Persistent_Value.xAutoEnabled
	AND (GVL_GEOMETRY_CONTROL.astStatus[1].xEnabled OR GVL_GEOMETRY_CONTROL.astStatus[2].xEnabled)
	AND (GVL_GEOMETRY_CONTROL.auiActiveCount[uiMachine] >= (MAX(UINT#1, Persistent_Value.auiPeriod[uiMachine]) - UINT#1)) THEN
		xCalled := TRUE;
	END_IF;
	xReadyDetail := astMachineStatus[uiMachine].xEnabled
		AND NOT astMachineStatus[uiMachine].xError AND NOT astMachineStatus[uiMachine].xDisablePending
		AND NOT astMachineStatus[uiMachine].xBusy AND NOT astMachineStatus[uiMachine].xProcessing
		AND astMachineStatus[uiMachine].xCanAcceptService AND astMachineStatus[uiMachine].xServiceRequired
		AND (astMachineStatus[uiMachine].ePartState = E_PART_STATE.LOADED)
		AND (astMachineStatus[uiMachine].ePartType = E_PART_TYPE.DETAIL);
	IF xRunning AND NOT xManual AND xCalled AND xReadyDetail AND (uiCallState <> UINT#1) THEN
		Persistent_Value.udiNextCallId := Persistent_Value.udiNextCallId + UDINT#1;
		IF Persistent_Value.udiNextCallId = UDINT#0 THEN Persistent_Value.udiNextCallId := UDINT#1; END_IF;
		Call := EmptyCall; Call.udiId := Persistent_Value.udiNextCallId;
		Call.uiMachine := uiMachine; Call.uiProductType := Config.auiMachineType[uiMachine]; Call.uiState := UINT#1;
		GVL_GEOMETRY_CONTROL.astCalls[uiMachine] := Call;
		F_GEOMETRY_EVENT(Call := Call);
	END_IF;
	// Пустой станок можно загрузить. Уже начатый рецепт не прерываем.
	axGeometryUnloadBlocked[uiMachine] := xCalled AND (uiFreeStation = UINT#0)
		AND (astMachineStatus[uiMachine].ePartState = E_PART_STATE.LOADED)
		AND NOT astMachineStatus[uiMachine].xBusy;
END_FOR;

// Возраст вызова не ограничивает обслуживание; ждём только свободного ГК.
FOR uiMachine := FIRST_MACHINE TO LAST_MACHINE DO
	xReadyDetail := astMachineStatus[uiMachine].xEnabled
		AND NOT astMachineStatus[uiMachine].xError AND NOT astMachineStatus[uiMachine].xDisablePending
		AND NOT astMachineStatus[uiMachine].xBusy AND NOT astMachineStatus[uiMachine].xProcessing
		AND astMachineStatus[uiMachine].xCanAcceptService AND astMachineStatus[uiMachine].xServiceRequired
		AND (astMachineStatus[uiMachine].ePartState = E_PART_STATE.LOADED)
		AND (astMachineStatus[uiMachine].ePartType = E_PART_TYPE.DETAIL);
	// W52 относится только к готовой детали без доступного свободного ГК.
	xWaiting := xRunning AND NOT xManual AND NOT xGlobalError
		AND xReadyDetail AND axGeometryUnloadBlocked[uiMachine] AND (uiFreeStation = UINT#0);
	// Отдельный TON для каждого вызова; реальное время, без ускорения симуляции.
	atonGeometryWait[uiMachine](IN := xWaiting AND NOT GVL_ALARM.Command.xResetWarnings
		AND (audiGeometryWaitCallId[uiMachine] = GVL_GEOMETRY_CONTROL.astCalls[uiMachine].udiId),
		PT := Persistent_Value.tWaitWarningTimeout);
	IF NOT xWaiting OR GVL_ALARM.Command.xResetWarnings
	OR (audiGeometryWaitCallId[uiMachine] <> GVL_GEOMETRY_CONTROL.astCalls[uiMachine].udiId) THEN
		axGeometryWaitWarned[uiMachine] := FALSE;
	END_IF;
	audiGeometryWaitCallId[uiMachine] := GVL_GEOMETRY_CONTROL.astCalls[uiMachine].udiId;
	IF atonGeometryWait[uiMachine].Q AND NOT axGeometryWaitWarned[uiMachine] THEN
		axGeometryWaitWarned[uiMachine] := TRUE; xRaiseWarning := TRUE;
	END_IF;
END_FOR;
IF xRaiseWarning THEN
	GVL_GEOMETRY_CONTROL.stCellWarning.uiCode := WRN_GEOMETRY_WAIT_TIMEOUT; // WARNING: остальные станки продолжают работу
	GVL_GEOMETRY_CONTROL.stCellWarning.udiSequence := GVL_GEOMETRY_CONTROL.stCellWarning.udiSequence + UDINT#1;
	IF GVL_GEOMETRY_CONTROL.stCellWarning.udiSequence = UDINT#0 THEN GVL_GEOMETRY_CONTROL.stCellWarning.udiSequence := UDINT#1; END_IF;
END_IF;
